FUNCTION_BLOCK E_DEMUX_FIFO_2 (* Gegenstueck zu E_MUX_FIFO_2_Adapter: verteilt DATA vom Socket IN_DATA nach dem Kanal (OUT = 0/1) auf EO1/EO2. PROCESSED vom Konsumenten geht ueber den Rueckkanal des Adapters zurueck, erst dann folgt das naechste Ereignis. *)
  (* Standard: 61499-2; Description: Copyright (c) 2026 Meisterschulen am Ostbahnhof This program and the accompanying materials are made available under the terms of the Eclipse Public License 2.0 which is available at https://www.eclipse.org/legal/epl-2.0/ SPDX-License-Identifier: EPL-2.0 *)
  (* Version 1.0, 2026-11-11, Franz Höpfinger, Meisterschulen am Ostbahnhof, initial API and implementation and/or initial documentation *)
  PACKAGE FIFO_adapter;
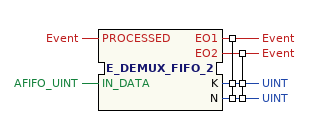
  EVENT_INPUT
    PROCESSED; (* Konsument bestaetigt: das zuletzt ausgegebene Ereignis ist verarbeitet *)
  END_EVENT
  EVENT_OUTPUT
    EO1 WITH K, N; (* Ereignis von Kanal 1 (K = 0) *)
    EO2 WITH K, N; (* Ereignis von Kanal 2 (K = 1) *)
  END_EVENT
  VAR_OUTPUT
    K : UINT; (* Kanal des ausgegebenen Ereignisses *)
    N : UINT; (* Anzahl der danach noch wartenden Ereignisse in der Queue *)
  END_VAR
  SOCKETS
    IN_DATA : FIFO_adapter::AFIFO_UINT; (* Hier haengt der Plug OUT_DATA von E_MUX_FIFO_2_Adapter an *)
  END_SOCKETS
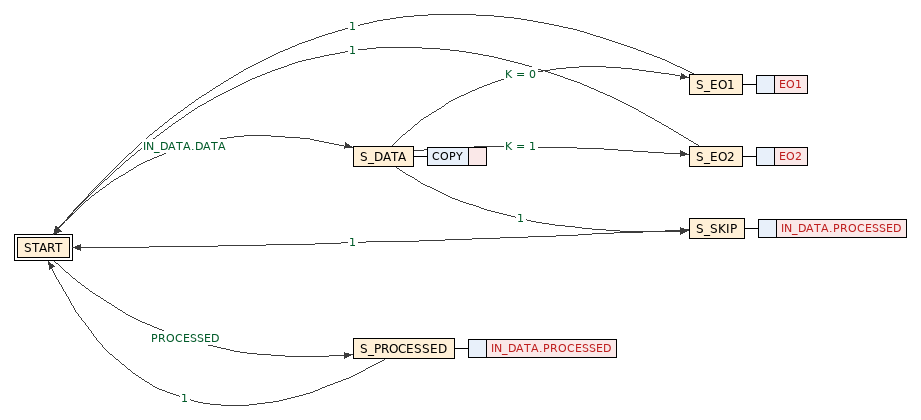
  EC_STATES
    START; (* Initial State *)
    S_DATA : COPY;
    S_EO1 : -> EO1;
    S_EO2 : -> EO2;
    S_SKIP : -> IN_DATA.PROCESSED; (* Unbekannter Kanal: sofort quittieren, sonst haengt die Queue *)
    S_PROCESSED : -> IN_DATA.PROCESSED;
  END_STATES
  EC_TRANSITIONS
    START TO S_DATA := IN_DATA.DATA;
    S_DATA TO S_EO1 := K = 0;
    S_DATA TO S_EO2 := K = 1;
    S_DATA TO S_SKIP := 1;
    S_EO1 TO START := 1;
    S_EO2 TO START := 1;
    S_SKIP TO START := 1;
    START TO S_PROCESSED := PROCESSED;
    S_PROCESSED TO START := 1;
  END_TRANSITIONS
  ALGORITHM COPY IN ST: (* Kanal und Fuellstand vom Adapter uebernehmen *)
K := IN_DATA.OUT;
N := IN_DATA.N;
  END_ALGORITHM
END_FUNCTION_BLOCK
